TYPE "ST_MeasRecord"
VERSION : 0.1
   STRUCT
      "Name" : String[64];
      "Value" : LReal;
      "Minimum" : LReal;
      "Maximum" : LReal;
      "Target" : LReal;
      "Unit" : String[16];
      "InTol" : Bool;
   END_STRUCT;
END_TYPE
